(* IEC 61131-3 sources: llm-plc-st-eval/data/raw/claude-sonnet-4-6/I1/few_shot, 3 files *)

(* ---- ejec_1.st ---- *)
```st
FUNCTION_BLOCK FB_Semaforo
VAR_INPUT
    habilitado : BOOL; (* Habilita la secuencia normal del semaforo *)
END_VAR
VAR_OUTPUT
    luzV : BOOL; (* Luz verde *)
    luzA : BOOL; (* Luz amarilla *)
    luzR : BOOL; (* Luz roja *)
END_VAR
VAR
    estado     : INT;  (* Estado actual: 0=Verde, 1=Amarillo, 2=Rojo, 3=Amarillo intermitente *)
    tFase      : TON; (* Temporizador de fase normal *)
    tBlink     : TP;  (* Temporizador de pulso para amarillo intermitente *)
    blinkCiclo : BOOL; (* Disparo ciclico del parpadeo *)
END_VAR

IF NOT habilitado THEN
    (* --- Modo amarillo intermitente --- *)
    estado := 3;

    (* Genera ciclos de 1 s usando TP: cuando Q baja, se relanza *)
    tBlink(IN := NOT tBlink.Q AND NOT blinkCiclo, PT := T#1S);

    (* blinkCiclo alterna cada vez que el temporizador termina *)
    IF tBlink.Q THEN
        blinkCiclo := NOT blinkCiclo;
    END_IF;

    luzV := FALSE;
    luzA := blinkCiclo; (* Amarillo parpadea 1 s ON / 1 s OFF *)
    luzR := FALSE;

    (* Reinicia el temporizador de fase para que al habilitar empiece limpio *)
    tFase(IN := FALSE, PT := T#1S);

ELSE
    (* --- Modo secuencia normal --- *)
    tBlink(IN := FALSE, PT := T#1S); (* Mantiene el TP inactivo *)
    blinkCiclo := FALSE;

    CASE estado OF

        0: (* Verde 20 s *)
            luzV := TRUE;
            luzA := FALSE;
            luzR := FALSE;
            tFase(IN := TRUE, PT := T#20S);
            IF tFase.Q THEN
                tFase(IN := FALSE, PT := T#20S); (* Resetea temporizador *)
                estado := 1;
            END_IF;

        1: (* Amarillo 4 s *)
            luzV := FALSE;
            luzA := TRUE;
            luzR := FALSE;
            tFase(IN := TRUE, PT := T#4S);
            IF tFase.Q THEN
                tFase(IN := FALSE, PT := T#4S);
                estado := 2;
            END_IF;

        2: (* Rojo 15 s *)
            luzV := FALSE;
            luzA := FALSE;
            luzR := TRUE;
            tFase(IN := TRUE, PT := T#15S);
            IF tFase.Q THEN
                tFase(IN := FALSE, PT := T#15S);
                estado := 0; (* Reinicia ciclo *)
            END_IF;

        3: (* Venia de modo intermitente: reinicia en verde *)
            estado := 0;
            tFase(IN := FALSE, PT := T#1S);
            luzV := FALSE;
            luzA := FALSE;
            luzR := FALSE;

        ELSE
            estado := 0; (* Estado invalido: ir a verde *)

    END_CASE;
END_IF;

END_FUNCTION_BLOCK
```

(* ---- ejec_2.st ---- *)
```st
FUNCTION_BLOCK FB_Semaforo
VAR_INPUT
    habilitado : BOOL; (* Habilitacion del semaforo *)
END_VAR
VAR_OUTPUT
    luzV : BOOL; (* Luz verde *)
    luzA : BOOL; (* Luz amarilla *)
    luzR : BOOL; (* Luz roja *)
END_VAR
VAR
    estado     : INT;  (* 0=Verde, 1=Amarillo, 2=Rojo, 3=Amarillo intermitente *)
    tFase      : TON; (* Temporizador de fase normal *)
    tBlink     : TP;  (* Temporizador de pulso para intermitente *)
    blinkState : BOOL; (* Estado actual del parpadeo *)
END_VAR

(* --- Maquina de estados del semaforo --- *)

IF NOT habilitado THEN
    (* Modo amarillo intermitente: las demas luces apagadas *)
    estado := 3;
    tFase(IN := FALSE, PT := T#1S); (* Resetear temporizador de fase *)
END_IF

CASE estado OF

    0: (* VERDE - 20 segundos *)
        luzV := TRUE;
        luzA := FALSE;
        luzR := FALSE;
        tFase(IN := TRUE, PT := T#20S);
        IF tFase.Q THEN
            tFase(IN := FALSE, PT := T#20S); (* Reset temporizador *)
            estado := 1;
        END_IF

    1: (* AMARILLO - 4 segundos *)
        luzV := FALSE;
        luzA := TRUE;
        luzR := FALSE;
        tFase(IN := TRUE, PT := T#4S);
        IF tFase.Q THEN
            tFase(IN := FALSE, PT := T#4S); (* Reset temporizador *)
            estado := 2;
        END_IF

    2: (* ROJO - 15 segundos *)
        luzV := FALSE;
        luzA := FALSE;
        luzR := TRUE;
        tFase(IN := TRUE, PT := T#15S);
        IF tFase.Q THEN
            tFase(IN := FALSE, PT := T#15S); (* Reset temporizador *)
            estado := 0; (* Reinicia ciclo en verde *)
        END_IF

    3: (* AMARILLO INTERMITENTE - 1s ON / 1s OFF *)
        luzV := FALSE;
        luzR := FALSE;
        (* Pulso de 1 segundo para generar el parpadeo *)
        tBlink(IN := NOT tBlink.Q, PT := T#1S);
        IF tBlink.Q THEN
            blinkState := NOT blinkState; (* Alternar estado del parpadeo *)
        END_IF
        luzA := blinkState;
        (* Si se habilita de nuevo, reiniciar en verde *)
        IF habilitado THEN
            blinkState := FALSE;
            tBlink(IN := FALSE, PT := T#1S); (* Reset temporizador blink *)
            estado := 0;
        END_IF

    ELSE
        (* Estado desconocido: ir a verde por seguridad *)
        estado := 0;

END_CASE

END_FUNCTION_BLOCK
```

(* ---- ejec_3.st ---- *)
```st
FUNCTION_BLOCK FB_Semaforo
VAR_INPUT
    habilitado : BOOL; (* Habilitacion del semaforo *)
END_VAR
VAR_OUTPUT
    luzV : BOOL; (* Luz verde *)
    luzA : BOOL; (* Luz amarilla *)
    luzR : BOOL; (* Luz roja *)
END_VAR
VAR
    estado     : INT;  (* Estado de la secuencia: 0=Verde, 1=Amarillo, 2=Rojo *)
    tFase      : TON; (* Temporizador de fase normal *)
    tBlink     : TP;  (* Temporizador de pulso para amarillo intermitente *)
    blinkState : BOOL; (* Estado actual del parpadeo (ON/OFF) *)
END_VAR

IF NOT habilitado THEN
    (* --- Modo amarillo intermitente --- *)
    estado := 0; (* Reinicio de estado para cuando se habilite de nuevo *)
    luzV   := FALSE;
    luzR   := FALSE;

    (* Generar parpadeo: cada flanco de bajada de tBlink.Q relanza el pulso *)
    tBlink(IN := NOT tBlink.Q, PT := T#1S);
    blinkState := tBlink.Q;
    luzA := blinkState;

    (* Asegurar que el temporizador de fase no quede activo *)
    tFase(IN := FALSE, PT := T#20S);

ELSE
    (* --- Modo secuencia normal --- *)
    tBlink(IN := FALSE, PT := T#1S); (* Detener y resetear el temporizador de parpadeo *)
    blinkState := FALSE;

    CASE estado OF

        0: (* Verde: 20 segundos *)
            luzV := TRUE;
            luzA := FALSE;
            luzR := FALSE;
            tFase(IN := TRUE, PT := T#20S);
            IF tFase.Q THEN
                tFase(IN := FALSE, PT := T#20S); (* Reset temporizador *)
                estado := 1;
            END_IF;

        1: (* Amarillo: 4 segundos *)
            luzV := FALSE;
            luzA := TRUE;
            luzR := FALSE;
            tFase(IN := TRUE, PT := T#4S);
            IF tFase.Q THEN
                tFase(IN := FALSE, PT := T#4S); (* Reset temporizador *)
                estado := 2;
            END_IF;

        2: (* Rojo: 15 segundos *)
            luzV := FALSE;
            luzA := FALSE;
            luzR := TRUE;
            tFase(IN := TRUE, PT := T#15S);
            IF tFase.Q THEN
                tFase(IN := FALSE, PT := T#15S); (* Reset temporizador *)
                estado := 0; (* Reinicia la secuencia *)
            END_IF;

        ELSE
            estado := 0; (* Estado invalido: volver a verde *)

    END_CASE;

END_IF;

END_FUNCTION_BLOCK
```
